FUNCTION f_QueuePop : BOOL
VAR_INPUT
    pQueue : POINTER TO T_StringQueue;
END_VAR
VAR_OUTPUT
    str : STRING(255);
END_VAR

IF pQueue^.Count <= 0 THEN
    f_QueuePop := FALSE; // Empty
ELSE
    str := pQueue^.Buffer[pQueue^.Head];
    pQueue^.Head := (pQueue^.Head + 1) MOD 20;
    pQueue^.Count := pQueue^.Count - 1;
    f_QueuePop := TRUE;
END_IF

END_FUNCTION

(* stored: Version 1.1.0.1, ProductVersion 3.1.4024.15
   POU f_QueuePop: Id {7ef47e54-316e-4974-affc-18f3f7a92706}, SpecialFunc None *)
